Staubli VAL3: utText.pjx

--- utText.pjx ---
Parameters version=s8.8.3Cs9_BS1660 stackSize=5000 millimeterUnit=true
Program file=start.pgx
Program file=stop.pgx
Data file=utText.dtx

--- utText.dtx ---
public string sFontFamily
public string sFontStyle
public string sFontWeight
public string sTextAlignment
public num nFontSize

--- start.pgx ---
program start()
begin
end

--- stop.pgx ---
program stop()
begin
end
